// TIA Portal V21 export
// export: Created 2026-11-22T02:34:46.634863Z, ExportSetting WithDefaults, DisplayName Totally Integrated Automation Portal, DisplayVersion V21 Update 3, DisplayName STEP 7 Professional, DisplayVersion V21 Update 3, DisplayName STEP 7 Safety, DisplayVersion V21, DisplayName Tech WebApplication, DisplayVersion V21, DisplayName WinCC Basic/Comfort/Advanced, DisplayVersion V21 Update 3, DisplayName WinCC Unified, DisplayVersion V21 Update 3
Screen "D_Gauge_2"  1024x768, Number=486
  ScreenLayer "Layer_0"
    Gauge "PV_Pct_MaxMin" at 6,4 size 150x150  CenterSize=0.08, DialSize=0.87, Gradation=10, InnerDialInnerDistance=0.08, InnerDialOuterDistance=0.9, MaximumValue=100, RangeUpper1Start=3.5, RangeUpper2Start=70, StyleItem=Gauge, CaptionText="SIMATIC"
      ProcessValue := D_Pct
      MaximumValue := D_Max
      MinimumValue := D_Min
    TextField "Label_PV_Pct_MaxMin" at 6,186 size 198x16  StyleItem=Text field, Text="PV_Pct_MaxMin"
    IOField "State" at 4,742 size 60x22  DataFormat=Decimal, FormatPattern=9, Mode=Output, StyleItem=I/O field
      ProcessValue := D_State
    Button "S1" at 70,742 size 40x22  Mode=Text, StyleItem=Button, TextOff="S1", TextOn="S1"
      on Click: SetS1()
    Button "S2" at 114,742 size 40x22  Mode=Text, StyleItem=Button, TextOff="S2", TextOn="S2"
      on Click: SetS2()
    Button "S3" at 158,742 size 40x22  Mode=Text, StyleItem=Button, TextOff="S3", TextOn="S3"
      on Click: SetS3()
    Button "S4" at 202,742 size 40x22  Mode=Text, StyleItem=Button, TextOff="S4", TextOn="S4"
      on Click: SetS4()
    Button "Next" at 980,742 size 40x22  Mode=Text, StyleItem=Button, TextOff="Next", TextOn="Next"
      on Click: ActivateScreen(Screen name := D_Clock_1, Object number := 0)
